(*
SPDX-FileCopyrightText: c 2026 Oleksandr Tiutyk <trofimich@gmail.com>
SPDX-License-Identifier: MIT
License: https://opensource.org/license/mit
*)

(*!
<summary>Checks input inversion for a normally closed contact.</summary>
<description>
Uses a live case-owned automation parent and fresh local device fixtures on every run.
The scenario reads and writes ordinary simulated storage within one task cycle.
</description>
*)

{attribute 'no_assign'}
{attribute 'no_explicit_call' := 'do not call this function block directly'}
FUNCTION_BLOCK DigitalInputNormallyClosedTest EXTENDS TOF_Testing.SingleCycleTest
VAR_STAT
	{attribute 'hide'}
	_ClassName : STRING := __POUNAME();
END_VAR
VAR
	//! <summary>Live parent borrowed by the method-local simulated device.</summary>
	_AutomationRoot : MockAutomationController(name := "DevicesIORoot");
END_VAR

(*!
<summary>Checks input inversion for a normally closed contact.</summary>
*)
METHOD PROTECTED ExecuteTest
VAR
	input : TOF_Devices_IO.DigitalInput(name := "DI_NC", parent := _AutomationRoot);
	rawInput : BOOL;
END_VAR
input.Initialize();
input.ContactType := TOF_Devices_IO.CONTACT_TYPE.NORMALLY_CLOSED;
input.BindToIO(rawValue := rawInput);

rawInput := FALSE;
input.ProcessInput();
Assert.ThatBool(
	actual := input.Value,
	message := "Value should be inverted TRUE for NC contact"
).IsTrue();

rawInput := TRUE;
input.ProcessInput();
Assert.ThatBool(
	actual := input.Value,
	message := "Value should be inverted FALSE for NC contact"
).IsFalse();
END_METHOD

//! <summary>Borrows the concrete class name. Callers must not modify it.</summary>
{attribute 'monitoring' := 'call'}
PROPERTY ClassName : REFERENCE TO STRING
GET
ClassName REF= _ClassName;
END_GET
END_PROPERTY

//! <summary>Borrows the compiler-initialized namespace name. Callers must not modify it.</summary>
{attribute 'monitoring' := 'call'}
PROPERTY NamespaceName : REFERENCE TO STRING
GET
NamespaceName REF= CurrentNamespace.Name;
END_GET
END_PROPERTY

//! <summary>Reports the concrete instance size in bytes.</summary>
{attribute 'monitoring' := 'call'}
PROPERTY SelfSize : ULINT
GET
SelfSize := XSIZEOF(THIS^);
END_GET
END_PROPERTY

END_FUNCTION_BLOCK

(* stored: Version 1.1.0.1
   POU DigitalInputNormallyClosedTest: Id {abee0954-0b0f-4551-b518-c01467414f49}, SpecialFunc None
   Method ExecuteTest: Id {c9ff93da-5480-4635-8a84-36bb1862c3d8}
   Property ClassName: Id {4c3d2a6c-cf35-43fa-9523-9da68990790f}
   Get Get: Id {f4b58111-a571-4052-af93-85a92a0aa28c}
   Property NamespaceName: Id {dd41f36c-e9d2-4503-8b17-8863b91b141a}
   Get Get: Id {a2474043-973c-4e10-995f-ab4e31f82096}
   Property SelfSize: Id {60ce3482-2ce0-49f6-b825-bff8a5c9a0db}
   Get Get: Id {e3bd5180-df3c-407b-b294-889afbf7aab4} *)
